TYPE ST_HmiCommands :
STRUCT
    bStart                 : BOOL;
    bStop                  : BOOL;
    bReset                 : BOOL;
    bAcknowledge           : BOOL;
    bManualRequest         : BOOL;
    bIndexerManualEnable   : BOOL;
    bManualIndexForward    : BOOL;
    bManualIndexHome       : BOOL;
    bManualMainDoorUnlock  : BOOL;
    uiResetStatisticsNestId: UINT;
END_STRUCT
END_TYPE

(* stored: Version 1.1.0.1, ProductVersion 3.1.4026.18
   DUT ST_HmiCommands: Id {cea0711c-b7bf-4958-9705-69290143acac} *)
